// Comparaison d'un terme de condition (docs/05 § 3.7)
{attribute 'qualified_only'}
{attribute 'strict'}
TYPE E_Cmp :
(
    Eq := 0,
    Ne := 1,
    Lt := 2,
    Le := 3,
    Gt := 4,
    Ge := 5,
    IsTrue := 6,
    IsFalse := 7
) USINT;
END_TYPE

(* stored: Version 1.1.0.1, ProductVersion 3.1.4024.12
   DUT E_Cmp: Id {0d90606f-5e55-523a-80c3-6891043d680b} *)
